(* IEC 61131-3 sources: BODAS-RC27-18_40/st/bodas_rc18_12_27_18_40/plc_logic/application/easyconfig_import/bds_syspb_ec, 2 files *)

(* ---- bds_syspb_vrnt_te-bds_sysPb_vrnt_te.st ---- *)
(* --- Interface --- *)
///post build system variants information
{attribute 'qualified_only' := ''}
{attribute 'strict' := ''}
TYPE bds_sysPb_vrnt_te :
(
	bds_sysPb_vrnt01_E  := 0,
	bds_sysPb_maxNumVrnt_E
) USINT;
END_TYPE

(* ---- bds_syspb_ec_gvl-bds_sysPb_ec_gvl.st ---- *)
(* --- Interface --- *)
{attribute 'qualified_only' := ''}
VAR_GLOBAL CONSTANT
	RC40: USINT := bds_sysPb_vrnt_te.bds_sysPb_vrnt01_E;
END_VAR
